{region 'Documentation'}
(*!
<summary>Named non-positive event publishing results; positive INT results indicate successful insertion.</summary>
*)
{endregion}
{attribute 'qualified_only'}
TYPE E_EventPublishResult : E_FifoResult;
END_TYPE

(* stored: Version 1.1.0.1
   DUT E_EventPublishResult: Id {8ad2cfb7-bfc7-491c-940c-e19d27885ee4} *)
